(* IEC 61131-3 sources: model-first-plc-agent-ai/gvm/generated, 1 file *)

(* ---- tank_reference_gvm.st ---- *)
(* Generated by gvm/grafcet2gvm.py from tank_reference.json (description SHA-256 278008e6fb70fcac); do not edit.
   GVM program: one tick = one evolution of the GRAFCET to a stable situation (semantics of
   nusmv/grafcet2smv.py, checked with NuSMV).
   Enumerated inputs as INT indices: mode: 0 timer, 1 tontof, 2 pid; r: 0 LOW, 1 MID, 2 HIGH.
   One scan of PROGRAM Main = one evolution; the situation is kept in the FB instance between scans. *)

FUNCTION_BLOCK FB_GVM_tank_reference
  VAR_INPUT
    in_start : BOOL;
    in_stop : BOOL;
    in_mode : INT;
    in_r : INT;
    in_timer_q : BOOL;
    in_ton_q : BOOL;
    in_tof_q : BOOL;
    in_hold_ok : BOOL;
    in_logged : BOOL;
  END_VAR
  VAR_OUTPUT
    out_fill_valve : BOOL;
    out_pid_on : BOOL;
    out_discharge_at_ud : BOOL;
    stable : BOOL;
    x0 : BOOL := TRUE;
    xE1 : BOOL := FALSE;
    xS1 : BOOL := FALSE;
    xE2 : BOOL := FALSE;
    x21 : BOOL := FALSE;
    x22 : BOOL := FALSE;
    xS2 : BOOL := FALSE;
    xE3 : BOOL := FALSE;
    xS3 : BOOL := FALSE;
    x4 : BOOL := FALSE;
    x5 : BOOL := FALSE;
    x6 : BOOL := FALSE;
    x10 : BOOL := TRUE;
    x11 : BOOL := FALSE;
  END_VAR
  VAR
    k_x0, k_xE1, k_xS1, k_xE2, k_x21, k_x22, k_xS2, k_xE3, k_xS3, k_x4, k_x5, k_x6, k_x10, k_x11 : BOOL;
    n_x0, n_xE1, n_xS1, n_xE2, n_x21, n_x22, n_xS2, n_xE3, n_xS3, n_x4, n_x5, n_x6, n_x10, n_x11 : BOOL;
    e_start, e_stop, e_timer_q, e_ton_q, e_tof_q, e_hold_ok, e_logged, d_LSH, d_LSHH, f_t0_E1, f_t0_E2, f_t0_E3, f_tE1_S1, f_tE2_21, f_t21_22, f_t21_S2, f_t22_21, f_tE3_S3, f_tEndM1, f_tEndM2, f_tEndM3, f_t4_56, f_t56_0, f_t10_11, f_t11_10 : BOOL;
    e_mode, e_r : INT;
    first : BOOL;
    m : INT;
  END_VAR
  k_x0 := x0;
  k_xE1 := xE1;
  k_xS1 := xS1;
  k_xE2 := xE2;
  k_x21 := x21;
  k_x22 := x22;
  k_xS2 := xS2;
  k_xE3 := xE3;
  k_xS3 := xS3;
  k_x4 := x4;
  k_x5 := x5;
  k_x6 := x6;
  k_x10 := x10;
  k_x11 := x11;
  FOR m := 1 TO 16 DO   (* K = 15 micro-steps, then one more for the stability check *)
    first := m = 1;
    IF first THEN e_start := in_start; ELSE e_start := FALSE; END_IF;
    e_stop := in_stop;
    e_mode := in_mode;
    e_r := in_r;
    IF k_xE1 THEN e_timer_q := in_timer_q; ELSE e_timer_q := FALSE; END_IF;
    IF k_x21 THEN e_ton_q := in_ton_q; ELSE e_ton_q := FALSE; END_IF;
    IF k_x22 THEN e_tof_q := in_tof_q; ELSE e_tof_q := TRUE; END_IF;
    IF k_xE3 THEN e_hold_ok := in_hold_ok; ELSE e_hold_ok := FALSE; END_IF;
    IF k_x6 THEN e_logged := in_logged; ELSE e_logged := FALSE; END_IF;
    d_LSH := ((e_r = 1) OR (e_r = 2));
    d_LSHH := (e_r = 2);
    f_t0_E1 := (x0 AND (e_start AND (e_mode = 0)));
    f_t0_E2 := (x0 AND (e_start AND (e_mode = 1)));
    f_t0_E3 := (x0 AND (e_start AND (e_mode = 2)));
    f_tE1_S1 := (xE1 AND (e_timer_q OR d_LSHH));
    f_tE2_21 := (xE2 AND TRUE);
    f_t21_22 := (x21 AND (e_ton_q AND NOT d_LSH));
    f_t21_S2 := (x21 AND d_LSH);
    f_t22_21 := (x22 AND NOT e_tof_q);
    f_tE3_S3 := (xE3 AND (e_hold_ok OR (e_r = 2)));
    f_tEndM1 := (xS1 AND TRUE);
    f_tEndM2 := (xS2 AND TRUE);
    f_tEndM3 := (xS3 AND TRUE);
    f_t4_56 := (x4 AND TRUE);
    f_t56_0 := ((x5 AND x6) AND e_logged);
    f_t10_11 := (x10 AND e_stop);
    f_t11_10 := (x11 AND NOT e_stop);
    n_x0 := ((x0 AND NOT ((f_t0_E1 OR f_t0_E2) OR f_t0_E3)) OR f_t56_0);
    n_xE1 := ((xE1 AND NOT f_tE1_S1) OR f_t0_E1);
    n_xS1 := ((xS1 AND NOT f_tEndM1) OR f_tE1_S1);
    n_xE2 := ((xE2 AND NOT f_tE2_21) OR f_t0_E2);
    n_x21 := ((x21 AND NOT (f_t21_22 OR f_t21_S2)) OR (f_tE2_21 OR f_t22_21));
    n_x22 := ((x22 AND NOT f_t22_21) OR f_t21_22);
    n_xS2 := ((xS2 AND NOT f_tEndM2) OR f_t21_S2);
    n_xE3 := ((xE3 AND NOT f_tE3_S3) OR f_t0_E3);
    n_xS3 := ((xS3 AND NOT f_tEndM3) OR f_tE3_S3);
    n_x4 := ((x4 AND NOT f_t4_56) OR ((f_tEndM1 OR f_tEndM2) OR f_tEndM3));
    n_x5 := ((x5 AND NOT f_t56_0) OR f_t4_56);
    n_x6 := ((x6 AND NOT f_t56_0) OR f_t4_56);
    n_x10 := ((x10 AND NOT f_t10_11) OR f_t11_10);
    n_x11 := ((x11 AND NOT f_t11_10) OR f_t10_11);
    IF n_x11 THEN
      n_x0 := TRUE;
      n_xE1 := FALSE;
      n_xS1 := FALSE;
      n_xE2 := FALSE;
      n_x21 := FALSE;
      n_x22 := FALSE;
      n_xS2 := FALSE;
      n_xE3 := FALSE;
      n_xS3 := FALSE;
      n_x4 := FALSE;
      n_x5 := FALSE;
      n_x6 := FALSE;
    END_IF;
    IF m <= 15 THEN
      k_x0 := k_x0 AND n_x0;
      k_xE1 := k_xE1 AND n_xE1;
      k_xS1 := k_xS1 AND n_xS1;
      k_xE2 := k_xE2 AND n_xE2;
      k_x21 := k_x21 AND n_x21;
      k_x22 := k_x22 AND n_x22;
      k_xS2 := k_xS2 AND n_xS2;
      k_xE3 := k_xE3 AND n_xE3;
      k_xS3 := k_xS3 AND n_xS3;
      k_x4 := k_x4 AND n_x4;
      k_x5 := k_x5 AND n_x5;
      k_x6 := k_x6 AND n_x6;
      k_x10 := k_x10 AND n_x10;
      k_x11 := k_x11 AND n_x11;
      x0 := n_x0;
      xE1 := n_xE1;
      xS1 := n_xS1;
      xE2 := n_xE2;
      x21 := n_x21;
      x22 := n_x22;
      xS2 := n_xS2;
      xE3 := n_xE3;
      xS3 := n_xS3;
      x4 := n_x4;
      x5 := n_x5;
      x6 := n_x6;
      x10 := n_x10;
      x11 := n_x11;
    ELSE
      stable := (n_x0 = x0) AND (n_xE1 = xE1) AND (n_xS1 = xS1) AND (n_xE2 = xE2) AND (n_x21 = x21) AND (n_x22 = x22) AND (n_xS2 = xS2) AND (n_xE3 = xE3) AND (n_xS3 = xS3) AND (n_x4 = x4) AND (n_x5 = x5) AND (n_x6 = x6) AND (n_x10 = x10) AND (n_x11 = x11);
    END_IF;
  END_FOR;
  out_fill_valve := ((xE1 OR x21) OR xE3);
  out_pid_on := xE3;
  out_discharge_at_ud := xE3;
END_FUNCTION_BLOCK

PROGRAM Main
  VAR
    pi_start AT %IX100.0 : BOOL;
    pi_stop AT %IX100.1 : BOOL;
    pi_mode AT %IW100 : INT;
    pi_r AT %IW101 : INT;
    pi_timer_q AT %IX100.2 : BOOL;
    pi_ton_q AT %IX100.3 : BOOL;
    pi_tof_q AT %IX100.4 : BOOL;
    pi_hold_ok AT %IX100.5 : BOOL;
    pi_logged AT %IX100.6 : BOOL;
    po_fill_valve AT %QX100.0 : BOOL;
    po_pid_on AT %QX100.1 : BOOL;
    po_discharge_at_ud AT %QX100.2 : BOOL;
    po_stable AT %QX100.3 : BOOL;
    px_x0 AT %QX101.0 : BOOL;
    px_xE1 AT %QX101.1 : BOOL;
    px_xS1 AT %QX101.2 : BOOL;
    px_xE2 AT %QX101.3 : BOOL;
    px_x21 AT %QX101.4 : BOOL;
    px_x22 AT %QX101.5 : BOOL;
    px_xS2 AT %QX101.6 : BOOL;
    px_xE3 AT %QX101.7 : BOOL;
    px_xS3 AT %QX102.0 : BOOL;
    px_x4 AT %QX102.1 : BOOL;
    px_x5 AT %QX102.2 : BOOL;
    px_x6 AT %QX102.3 : BOOL;
    px_x10 AT %QX102.4 : BOOL;
    px_x11 AT %QX102.5 : BOOL;
  END_VAR
  VAR
    gvm : FB_GVM_tank_reference;
  END_VAR
  gvm(in_start := pi_start, in_stop := pi_stop, in_mode := pi_mode, in_r := pi_r, in_timer_q := pi_timer_q, in_ton_q := pi_ton_q, in_tof_q := pi_tof_q, in_hold_ok := pi_hold_ok, in_logged := pi_logged);
  po_fill_valve := gvm.out_fill_valve;
  po_pid_on := gvm.out_pid_on;
  po_discharge_at_ud := gvm.out_discharge_at_ud;
  po_stable := gvm.stable;
  px_x0 := gvm.x0;
  px_xE1 := gvm.xE1;
  px_xS1 := gvm.xS1;
  px_xE2 := gvm.xE2;
  px_x21 := gvm.x21;
  px_x22 := gvm.x22;
  px_xS2 := gvm.xS2;
  px_xE3 := gvm.xE3;
  px_xS3 := gvm.xS3;
  px_x4 := gvm.x4;
  px_x5 := gvm.x5;
  px_x6 := gvm.x6;
  px_x10 := gvm.x10;
  px_x11 := gvm.x11;
END_PROGRAM
